Staubli VAL3: saveData.dtx

public bool bMarked
frame fMFrame = {fatherId=world[0]}
public frameItem fFrameItem[11]
  [0]
    frame fFrame = {fatherId=world[0]}
    pointRx pPointRx[3]
      [0] = {fatherId=world[0]}
      [1] = {fatherId=world[0]}
      [2] = {fatherId=world[0]}
    string sName = "world"
  [1]
    frame fFrame = {x=11, fatherId=world[0]}
    pointRx pPointRx[3]
      [0] = {x=490.0617294, y=-117.398102, z=1260.317878, rx=11.00784132, ry=17.654342, rz=-7.498705, shoulder=lefty, elbow=enegative, wrist=wpositive, fatherId=world[0]}
      [1] = {x=531.0703141, y=-117.398383, z=1260.317007, rx=11.00694015, ry=17.654895, rz=-7.49844, shoulder=lefty, elbow=enegative, wrist=wpositive, fatherId=world[0]}
      [2] = {x=531.0263881, y=-87.685862, z=1260.317101, rx=11.00680531, ry=17.654897, rz=-7.498382, shoulder=lefty, elbow=enegative, wrist=wpositive, fatherId=world[0]}
    string sName = "frame1"
  [2]
    frame fFrame = {x=574.25189, y=-115.239268, z=20.0712124, rx=0.00000547002, ry=0.0000199817, rz=0.0000210035, fatherId=world[0]}
    pointRx pPointRx[3]
      [0] = {x=574.25189, y=-115.239268, z=20.0712124, rx=3.180184, ry=-178.774731, rz=1.00275497, shoulder=lefty, elbow=epositive, wrist=wpositive, fatherId=world[0]}
      [1] = {x=713.860198, y=-115.239216, z=20.0711637, rx=3.179917, ry=-178.775635, rz=1.00265398, shoulder=lefty, elbow=epositive, wrist=wpositive, fatherId=world[0]}
      [2] = {x=713.810457, y=248.363282, z=20.0711985, rx=3.180844, ry=-178.775032, rz=1.0022136, shoulder=lefty, elbow=epositive, wrist=wpositive, fatherId=world[0]}
    string sName = "frame2"
  [3]
    frame fFrame = {fatherId=world[0]}
    pointRx pPointRx[3]
      [0] = {fatherId=world[0]}
      [1] = {fatherId=world[0]}
      [2] = {fatherId=world[0]}
    string sName = "frame3"
  [4]
    frame fFrame = {fatherId=world[0]}
    pointRx pPointRx[3]
      [0] = {fatherId=world[0]}
      [1] = {fatherId=world[0]}
      [2] = {fatherId=world[0]}
    string sName = "frame4"
  [5]
    frame fFrame = {fatherId=world[0]}
    pointRx pPointRx[3]
      [0] = {fatherId=world[0]}
      [1] = {fatherId=world[0]}
      [2] = {fatherId=world[0]}
    string sName = "frame5"
  [6]
    frame fFrame = {fatherId=world[0]}
    pointRx pPointRx[3]
      [0] = {fatherId=world[0]}
      [1] = {fatherId=world[0]}
      [2] = {fatherId=world[0]}
    string sName = "frame6"
  [7]
    frame fFrame = {fatherId=world[0]}
    pointRx pPointRx[3]
      [0] = {fatherId=world[0]}
      [1] = {fatherId=world[0]}
      [2] = {fatherId=world[0]}
    string sName = "frame7"
  [8]
    frame fFrame = {fatherId=world[0]}
    pointRx pPointRx[3]
      [0] = {fatherId=world[0]}
      [1] = {fatherId=world[0]}
      [2] = {fatherId=world[0]}
    string sName = "frame8"
  [9]
    frame fFrame = {fatherId=world[0]}
    pointRx pPointRx[3]
      [0] = {fatherId=world[0]}
      [1] = {fatherId=world[0]}
      [2] = {fatherId=world[0]}
    string sName = "frame9"
  [10]
    frame fFrame = {fatherId=world[0]}
    pointRx pPointRx[3]
      [0] = {fatherId=world[0]}
      [1] = {fatherId=world[0]}
      [2] = {fatherId=world[0]}
    string sName = "frame10"
public jointRx jHome = {j1=-6.654137, j2=-3.724613, j3=129.0455616, j4=-6.346552, j5=-34.647483, j6=4.794664}
mdesc mNomSpeed
public num nJogTool = 1
public num nLibIndex
public num nMarkIndex
public num nUsingTool = 1
public num sUsingLib
public pointRx pPowerOFF = {fatherId=world[0]}
public pointRx pPowerON = {fatherId=world[0]}
tool tMTool = {y=-160, z=500, fatherId=flange[0]}
public tool tUsingTool = {fatherId=flange[0]}
public toolItem tToolItem[11]
  [0]
    string sName = "flange"
    tool tTool = {fatherId=flange[0]}
  [1]
    string sName = "maintool"
    tool tTool = {x=1160, z=70, ry=-90, fatherId=flange[0]}
  [2]
    string sName = "tool2"
    tool tTool = {fatherId=flange[0]}
  [3]
    string sName = "tool3"
    tool tTool = {fatherId=flange[0]}
  [4]
    string sName = "tool4"
    tool tTool = {fatherId=flange[0]}
  [5]
    string sName = "tool5"
    tool tTool = {fatherId=flange[0]}
  [6]
    string sName = "tool6"
    tool tTool = {fatherId=flange[0]}
  [7]
    string sName = "tool7"
    tool tTool = {fatherId=flange[0]}
  [8]
    string sName = "tool8"
    tool tTool = {fatherId=flange[0]}
  [9]
    string sName = "tool9"
    tool tTool = {fatherId=flange[0]}
  [10]
    string sName = "tool10"
    tool tTool = {fatherId=flange[0]}
